(* ================================================================= *)
(*  ST_ExternalDevice                                                 *)
(*  外部设备接口结构体 - 状态/业务/控制/报警 四段式                    *)
(*  版本: V1.0.0  日期: 2026-05-20                                    *)
(*  来源: SysLib/types/                                               *)
(*  复用: 组框机/打胶机/机器人等上下游设备交互                         *)
(* ================================================================= *)

TYPE ST_ExternalDevice :
STRUCT
    // === 状态输入 (BOOL) ===
    AutoRunning     : BOOL := FALSE;   // 自动运行中
    Fault           : BOOL := FALSE;   // 设备故障
    EStop           : BOOL := FALSE;   // 急停状态
    CommError       : BOOL := FALSE;   // 通讯异常

    // === 业务信号 (BOOL) ===
    AllowFeed       : BOOL := FALSE;   // 允许送料/允许抓料
    PickupComplete  : BOOL := FALSE;   // 取料完成/堆垛完成
    MaterialRequest : BOOL := FALSE;   // 有料请求

    // === 控制输出 (BOOL) ===
    RequestRun      : BOOL := FALSE;   // 请求运行
    Pause           : BOOL := FALSE;   // 暂停
    ResetReq        : BOOL := FALSE;   // 复位请求
    Ready           : BOOL := FALSE;   // 本机就绪通知

    // === 报警汇总 (INT) ===
    DeviceAlarmCode : INT := 0;        // 设备专用报警码 (300~399)
END_STRUCT
END_TYPE
